Yaskawa INFORM job: PRECPRO.JBI

/JOB
//NAME PRECPRO
//POS
///NPOS 6,0,6,0,0,0
///TOOL 9
///POSTYPE PULSE
///PULSE
C00000=0,0,0
C00001=0,0,0
C00002=0,0,0
C00003=0,0,0
C00004=0,0,0
C00005=0,0,0
EC00000=0
EC00001=0
EC00002=0
EC00003=0
EC00004=0
EC00005=0
//INST
<volatile>
///COMM Generated using RoboDK
///ATTR SC,RW
///GROUP1 RB1
NOP
'Program generated by RoboDK v
'6.0.7 for Yaskawa Motoman EPL
'160 on XX/XX/XXXX 18:00:00
'Using nominal kinematics.
'Using Frame P (targets wrt ba
'se):
'0.0,-0.0,1000.0,90.0,-0.5,0.1
'Tool Tool P should be close t
'o:
'0.1,-0.4,123.5,-45.2,0.0,0.0
MOVJ C00000 VJ=50.00  +MOVJ EC00000 VJ=100.00
MOVL C00001 V=100.0  +MOVJ EC00001 VJ=100.00
MOVL C00002 V=100.0  +MOVJ EC00002 VJ=100.00
MOVJ C00003 VJ=50.00  +MOVJ EC00003 VJ=100.00
MOVJ C00004 VJ=50.00  +MOVJ EC00004 VJ=100.00
TIMER T=0.00
TIMER T=1.00
MOVL C00005 V=66.7  +MOVJ EC00005 VJ=100.00
END
